PROGRAM main
  VAR
    CONVEYOR AT %QX0.1 : BOOL;
  END_VAR

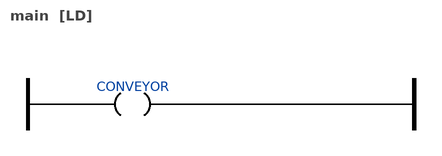
(* LD diagram, written out as Structured Text *)
CONVEYOR := TRUE;
END_PROGRAM
